(* IEC 61131-3 sources: bcs-engineering-dsl/language/test/generating/nested_control_test/expected, 4 files *)

(* ---- ProcessState.st ---- *)
{attribute 'qualified_only'}
{attribute 'strict'}
TYPE ProcessState :
(
    INIT := 0,
    PROCESSING := 1,
    FINALIZING := 2,
    COMPLETE := 3
);
END_TYPE

(* ---- NestedControlsFB_decl.st ---- *)
FUNCTION_BLOCK NestedControlsFB
VAR_INPUT
    iState: ProcessState;
    iCount: INT;
    iThreshold: REAL;
    iValues: ARRAY [0..9] OF REAL;
END_VAR
VAR_OUTPUT
    oResult: REAL;
    oStatus: STRING;
    oProcessedItems: INT;
END_VAR
VAR
    i: INT;
    tempSum: REAL := 0;
    itemsProcessed: INT := 0;
    skipCount: INT := 0;
END_VAR

(* ---- MAIN_decl.st ---- *)
PROGRAM MAIN
VAR
    TestNestedControls_state: ProcessState := ProcessState.PROCESSING;
    TestNestedControls_count: INT := 5;
    TestNestedControls_threshold: REAL := 10;
    TestNestedControls_values: ARRAY [0..9] OF REAL := [5, 15, 25, 7.5, 30, 0, 0, 0, 0, 0];
    TestNestedControls_result: REAL;
    TestNestedControls_status: STRING;
    TestNestedControls_processedItems: INT;
    NestedControlsFBInstance1: NestedControlsFB;
END_VAR

(* ---- NestedControlsFB_impl.st ---- *)
tempSum := 0;
itemsProcessed := 0;
skipCount := 0;
IF iState = ProcessState.INIT OR iState = ProcessState.PROCESSING THEN
    FOR i := 0 TO 9 BY 1 DO
        IF iValues[i] < iThreshold THEN
            skipCount := skipCount + 1;
            CONTINUE;
        END_IF;
        CASE iState OF
            ProcessState.INIT:
                tempSum := tempSum + iValues[i] * 0.8;
            ProcessState.PROCESSING:
                IF iValues[i] > iThreshold * 2 THEN
                    tempSum := tempSum + iValues[i] * 1.5;
                ELSE
                    tempSum := tempSum + iValues[i];
                END_IF;
            ELSE
                tempSum := tempSum + iValues[i] * 0.5;
        END_CASE;
        itemsProcessed := itemsProcessed + 1;
    END_FOR;
ELSIF iState = ProcessState.FINALIZING THEN
    tempSum := 0;
    i := 0;
    WHILE i < iCount AND i < 10 DO
        tempSum := tempSum + iValues[i] * 1.2;
        i := i + 1;
    END_WHILE;
    itemsProcessed := i;
ELSE
    tempSum := -1;
    itemsProcessed := 0;
END_IF;
oResult := tempSum;
oProcessedItems := itemsProcessed;
IF itemsProcessed = 0 THEN
    oStatus := 'No items processed';
ELSIF skipCount > 0 THEN
    oStatus := 'Processed with skips';
ELSE
    oStatus := 'All items processed';
END_IF;
